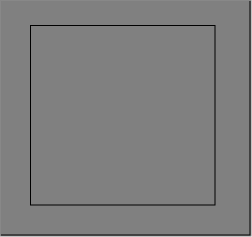
VISUALIZATION Sensor  // 252x237
VAR_INPUT
	{attribute 'parameterstringof' := 'm_Input_Sen_Addr'}
	m_Input_Sen_Addr_Str : STRING;
END_VAR
VAR_INPUT
	m_Input_Sen_Addr : Bool;
END_VAR
    Rectangle (0,0 250x235)
    RoundedRectangle (30,25 185x180), tooltip "%s", colour toggle: (m_Input_Sen_Addr) <> 0
        p4168582468: m_Input_Sen_Addr_Str
END_VISUALIZATION

(* stored: Version 1.1.0.1, ProductVersion 3.1.4024.13
   Visu Sensor: Id {397fc6ab-e589-4f3e-a401-78e81df10195} *)
